(* IEC 61131-3 sources: NachHouse_TST/TEST_Api/TEST_Api, 9 files *)

(* ---- 01_Types.st ---- *)
TYPE T_ROOM_CONFIG :
STRUCT
    Id              : USINT;
    Name            : STRING[32];
    ShortName       : STRING[12];
    FloorId         : USINT;
    SortOrder       : USINT;
    Icon            : STRING[24];
    Enabled         : BOOL;

    ShowTemperature : BOOL;
    ShowHumidity    : BOOL;
    ShowLights      : BOOL;
    ShowBlinds      : BOOL;
    ShowHeating     : BOOL;

    Image           : STRING[32];   // napr. livingroom.jpg
END_STRUCT
END_TYPE

TYPE T_ROOM_STATE :
STRUCT
    Temperature     : REAL;
    Humidity        : REAL;
    LightLevel      : UINT;

    LightsCount     : USINT;
    LightsOnCount   : USINT;
    LightsOn        : BOOL;

    BlindsCount     : USINT;
    BlindsMoving    : BOOL;
    BlindsPosition  : USINT;    // 0..100

    HeatingActive   : BOOL;
    CoolingActive   : BOOL;
    Setpoint        : REAL;

    AlarmActive     : BOOL;
    WarningActive   : BOOL;
    Occupied        : BOOL;

    ChangeCounter   : UDINT;
END_STRUCT
END_TYPE
(*
TYPE T_ROOM_CONFIG :
STRUCT
    Id          : USINT;
    Name        : STRING[32];
    ShortName   : STRING[12];
    FloorId     : USINT;
    SortOrder   : USINT;
    Icon        : STRING[24];
    Enabled     : BOOL;
END_STRUCT
END_TYPE

TYPE T_ROOM_STATE :
STRUCT
    Temperature     : REAL;
    Humidity        : REAL;
    LightLevel      : UINT;

    LightsCount     : USINT;
    LightsOnCount   : USINT;
    LightsOn        : BOOL;

    BlindsCount     : USINT;
    BlindsMoving    : BOOL;

    HeatingActive   : BOOL;
    CoolingActive   : BOOL;

    AlarmActive     : BOOL;
    WarningActive   : BOOL;
    Occupied        : BOOL;

    ChangeCounter   : UDINT;
END_STRUCT
END_TYPE
*)

TYPE T_API_CONFIG :
STRUCT
    Version         : UDINT;
    RoomCount       : USINT;
    Rooms           : ARRAY[1..8]   OF T_ROOM_CONFIG;
//    Lights          : ARRAY[1..300] OF T_LIGHT_CONFIG;
//    Blindss         : ARRAY[1..80]  OF T_BLIND_CONFIG;
//   ......
//   .....
END_STRUCT
END_TYPE

TYPE T_API_STATE :
STRUCT
    Version         : UDINT;
    Online          : BOOL;
    Counter         : UDINT;
    Rooms           : ARRAY[1..8] OF T_ROOM_STATE;
END_STRUCT
END_TYPE

TYPE T_API_COMMAND_REQUEST :
STRUCT
    RequestId       : UDINT;
    RoomId          : USINT;
    DeviceId        : UINT;
    Command         : USINT;

    ValueBool       : BOOL;
    ValueInt        : DINT;
    ValueReal       : REAL;

    Execute         : BOOL;
END_STRUCT
END_TYPE

TYPE T_API_COMMAND_RESULT :
STRUCT
    RequestId       : UDINT;
    ResultCode      : INT;
    Finished        : BOOL;
END_STRUCT
END_TYPE

TYPE T_API_COMMAND :
STRUCT
    Request         : T_API_COMMAND_REQUEST;
    Result          : T_API_COMMAND_RESULT;
END_STRUCT
END_TYPE

(* ---- 02_Constants.st ---- *)
VAR_GLOBAL CONSTANT
    C_ROOM_MAX : USINT := 8;

    CMD_NONE            : USINT := 0;
    CMD_ROOM_LIGHTS_OFF : USINT := 1;
    CMD_ROOM_LIGHTS_ON  : USINT := 2;

    RESULT_OK               : INT := 0;
    RESULT_UNKNOWN_COMMAND  : INT := -1;
    RESULT_INVALID_ROOM     : INT := -2;
    RESULT_INVALID_DEVICE   : INT := -3;
    RESULT_INVALID_VALUE    : INT := -4;
END_VAR

(* ---- 03_GVL_PublicApi.st ---- *)
VAR_GLOBAL
    ApiConfig {PUBLIC_API}  : T_API_CONFIG;
    ApiState   {PUBLIC_API} : T_API_STATE;
    ApiCommand  {PUBLIC_API} : T_API_COMMAND;
END_VAR

// new test var
VAR_GLOBAL
    TestWrite     {PUBLIC_API} : BOOL ;
//    MyTestApiVar1 {PUBLIC_API} : ARRAY[0..4] of STRING[255] ;
END_VAR

(* ---- 04_GVL_Internal.st ---- *)
VAR_GLOBAL
    ApiInitialized  : BOOL;
    LastRequestId   : UDINT;
END_VAR

(* ---- 05_prgApiInit.st ---- *)
FUNCTION prgApiInit : BOOL
VAR
    i : USINT;
END_VAR

IF NOT ApiInitialized THEN

    FOR i := 1 TO C_ROOM_MAX DO
        ApiConfig.Rooms[i].Id          := 0;
        ApiConfig.Rooms[i].Name        := '';
        ApiConfig.Rooms[i].ShortName   := '';
        ApiConfig.Rooms[i].FloorId     := 0;
        ApiConfig.Rooms[i].SortOrder   := 0;
        ApiConfig.Rooms[i].Icon        := '';
        ApiConfig.Rooms[i].Enabled     := FALSE;

        ApiState.Rooms[i].Temperature   := 0.0;
        ApiState.Rooms[i].Humidity      := 0.0;
        ApiState.Rooms[i].LightLevel    := 0;
        ApiState.Rooms[i].LightsCount   := 0;
        ApiState.Rooms[i].LightsOnCount := 0;
        ApiState.Rooms[i].LightsOn      := FALSE;
        ApiState.Rooms[i].BlindsCount   := 0;
        ApiState.Rooms[i].BlindsMoving  := FALSE;
        ApiState.Rooms[i].HeatingActive := FALSE;
        ApiState.Rooms[i].CoolingActive := FALSE;
        ApiState.Rooms[i].AlarmActive   := FALSE;
        ApiState.Rooms[i].WarningActive := FALSE;
        ApiState.Rooms[i].Occupied      := FALSE;
        ApiState.Rooms[i].ChangeCounter := 0;
    END_FOR;

    ApiConfig.Version   := 1;
    ApiConfig.RoomCount := 2;

    ApiConfig.Rooms[1].Id        := 1;
    ApiConfig.Rooms[1].Name      := 'Obyvacka';
    ApiConfig.Rooms[1].ShortName := 'Obyv.';
    ApiConfig.Rooms[1].FloorId   := 1;
    ApiConfig.Rooms[1].SortOrder := 1;
    ApiConfig.Rooms[1].Icon      := 'living_room';
    ApiConfig.Rooms[1].Enabled   := TRUE;

    ApiConfig.Rooms[2].Id        := 2;
    ApiConfig.Rooms[2].Name      := 'Kuchyna';
    ApiConfig.Rooms[2].ShortName := 'Kuch.';
    ApiConfig.Rooms[2].FloorId   := 1;
    ApiConfig.Rooms[2].SortOrder := 2;
    ApiConfig.Rooms[2].Icon      := 'kitchen';
    ApiConfig.Rooms[2].Enabled   := TRUE;

    ApiState.Version := 1;
    ApiState.Online  := TRUE;
    ApiState.Counter := 0;

    ApiState.Rooms[1].Temperature := 22.5;
    ApiState.Rooms[1].Humidity    := 45.0;
    ApiState.Rooms[1].LightLevel  := 350;
    ApiState.Rooms[1].LightsCount := 4;

    ApiState.Rooms[2].Temperature := 23.0;
    ApiState.Rooms[2].Humidity    := 48.0;
    ApiState.Rooms[2].LightLevel  := 250;
    ApiState.Rooms[2].LightsCount := 3;

    ApiCommand.Request.RequestId := 0;
    ApiCommand.Request.RoomId    := 0;
    ApiCommand.Request.DeviceId  := 0;
    ApiCommand.Request.Command   := CMD_NONE;
    ApiCommand.Request.ValueBool := FALSE;
    ApiCommand.Request.ValueInt  := 0;
    ApiCommand.Request.ValueReal := 0.0;
    ApiCommand.Request.Execute   := FALSE;

    ApiCommand.Result.RequestId  := 0;
    ApiCommand.Result.ResultCode := RESULT_OK;
    ApiCommand.Result.Finished   := FALSE;

    LastRequestId  := 0;
    ApiInitialized := TRUE;

END_IF;

END_FUNCTION

(* ---- 06_prgApiState.st ---- *)
FUNCTION prgApiState : BOOL
VAR
END_VAR

ApiState.Online  := TRUE;
// ApiState.Counter := ApiState.Counter + 1;

END_FUNCTION

(* ---- 07_prgApiCommand.st ---- *)
FUNCTION_BLOCK FBprgApiCommand
VAR
    RoomIndex : USINT;
END_VAR

IF ApiCommand.Request.Execute THEN

    IF ApiCommand.Request.RequestId <> LastRequestId THEN

        ApiCommand.Result.Finished   := FALSE;
        ApiCommand.Result.RequestId  := ApiCommand.Request.RequestId;
        ApiCommand.Result.ResultCode := RESULT_OK;

        RoomIndex := ApiCommand.Request.RoomId;

        IF (RoomIndex < 1) OR (RoomIndex > ApiConfig.RoomCount) THEN

            ApiCommand.Result.ResultCode := RESULT_INVALID_ROOM;

        ELSE

            CASE ApiCommand.Request.Command OF

                CMD_ROOM_LIGHTS_OFF:
                    ApiState.Rooms[RoomIndex].LightsOn      := FALSE;
                    ApiState.Rooms[RoomIndex].LightsOnCount := 0;
                    ApiState.Rooms[RoomIndex].ChangeCounter :=
                        ApiState.Rooms[RoomIndex].ChangeCounter + 1;

                CMD_ROOM_LIGHTS_ON:
                    ApiState.Rooms[RoomIndex].LightsOn := TRUE;
                    ApiState.Rooms[RoomIndex].LightsOnCount :=
                        ApiState.Rooms[RoomIndex].LightsCount;
                    ApiState.Rooms[RoomIndex].ChangeCounter :=
                        ApiState.Rooms[RoomIndex].ChangeCounter + 1;

                ELSE
                    ApiCommand.Result.ResultCode := RESULT_UNKNOWN_COMMAND;

            END_CASE;

        END_IF;

        LastRequestId := ApiCommand.Request.RequestId;
        ApiCommand.Result.Finished := TRUE;

    END_IF;

    ApiCommand.Request.Execute := FALSE;

END_IF;

END_FUNCTION_BLOCK

VAR_GLOBAL
   prgApiCommand : FBprgApiCommand;
END_VAR

(* ---- 08_MainProgram.st ---- *)
PROGRAM MainProgram
VAR
END_VAR

prgApiInit();
prgApiState();
prgApiCommand();

END_PROGRAM

(* ---- prgMain.ST ---- *)
PROGRAM prgMain
  VAR_INPUT
  END_VAR
  VAR_OUTPUT
  END_VAR
  VAR
  END_VAR
  VAR_TEMP
  END_VAR

   prgApiInit();
   prgApiState();
   prgApiCommand();

END_PROGRAM
